(* Logix 5000 project; controller TFF vendor 1 type 14 code 107 rev 33.11; software revision 33.04; part 28 of 38 *)
(* tags used below, declared in another part *)
   Address : DINT;   // Temp Address
   AO1 : ALIAS FOR AnalogOutput[8];
   AO2 : ALIAS FOR AnalogOutput[9];
   AO3 : ALIAS FOR AnalogOutput[10];
   AO4 : ALIAS FOR AnalogOutput[11];
   ControlLoop_FeedBagLevel : ALIAS FOR ControlLoop[2];
   ControlLoop_FeedBagLevelAlarm : ALIAS FOR AlarmDeviation[2];
   DF48MIX : ALIAS FOR DigitalPoint[26];
   DF48P001 : ALIAS FOR DigitalPoint[23];
   DF48P002 : ALIAS FOR DigitalPoint[24];
   DigitalOutput : BOOL[256];   // Digital Output Array these bits are sent to output cards.
   DigitalPoint : DigitalPoint[150];   // Digital Point Array
   DO1 : ALIAS FOR DigitalOutput[80];
   DO2 : ALIAS FOR DigitalOutput[81];
   DO3 : ALIAS FOR DigitalOutput[82];
   DO4 : ALIAS FOR DigitalOutput[83];
   DO5 : ALIAS FOR DigitalOutput[84];
   DO6 : ALIAS FOR DigitalOutput[85];
   DO7 : ALIAS FOR DigitalOutput[86];
   Drive : Drive[11];   // Drives Array
   Exchange_OUT : Exchange_OUT;   // Exchange Outputs
   FlowPath : FlowPath[64];   // Flow Path Array
   MIX101DF : ALIAS FOR DigitalPoint[28];
   Mixer : Mixer;   // Mixer config. structure
   Options : Options;   // Options List
   Phase0 : ALIAS FOR Phase[0];   // Phase 0
   PI401 : ALIAS FOR AnalogPoint[8];
   PipeAnimation : PipeAnimation;   // HMI Pipe Animation Array
   SIC001DF : ALIAS FOR DigitalPoint[16];
   SIC002 : ALIAS FOR Drive[2];
   SIC002DF : ALIAS FOR DigitalPoint[17];
   SIC004 : ALIAS FOR Drive[3];
   SysControl : SysControl;   // General system status and command
   Tank : TankManagement;   // Tank Management
   WI101 : ALIAS FOR AnalogPoint[15];
(* Process, continued *)

ROUTINE Drive_SIC002_Transfer   (* ladder *)
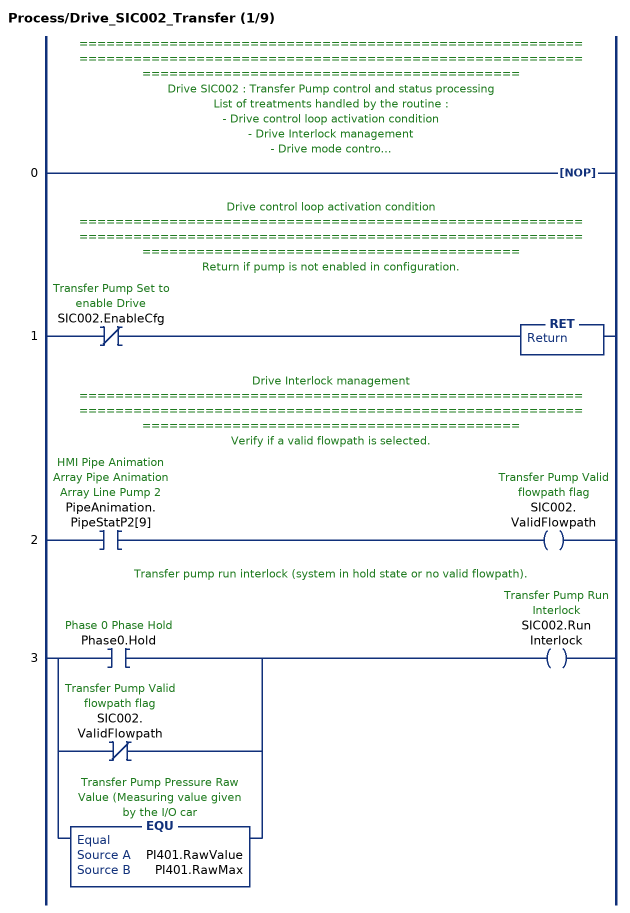
   // ==========================================================================================================================================================
   //                                                              Drive SIC002 : Transfer Pump control and status processing
   //                                                     List of treatments handled by the routine :
   //                                                          - Drive control loop activation condition
   //                                                          - Drive Interlock management
   //                                                          - Drive mode control
   //                                                          - Drive run command control
   //                                                          - Drive status management
   //                                                          - Drive status for HMI
   //                                                          - Drive DigitalOutput control
   //                                                     -----------------------------------------------------------------------------------------------------------------------------------------------------
   //                                                     History
   // 		2019-DEC-24 - Merck - Q. Spindler - Initial version for Candidate Release 1.00.00.00.a
   // 		2020-APR-06 - Merck - Q. Spindler - Modifications for Candidate Release 1.00.00.00.b
   //                                                                     - Add interlock when PI401 raw value is equal to RawMax (Sensor disconected)
   // ==========================================================================================================================================================
   0: NOP();
   // Drive control loop activation condition
   // ==========================================================================================================================================================
   // Return if pump is not enabled in configuration.
   1: XIO(SIC002.EnableCfg)RET();
   // Drive Interlock management
   // ==========================================================================================================================================================
   // Verify if a valid flowpath is selected.
   2: XIC(PipeAnimation.PipeStatP2[9])OTE(SIC002.ValidFlowpath);
   // Transfer pump run interlock (system in hold state or no valid flowpath).
   3: [XIC(Phase0.Hold) ,XIO(SIC002.ValidFlowpath) ,EQU(PI401.RawValue,PI401.RawMax) ]OTE(SIC002.RunInterlock);
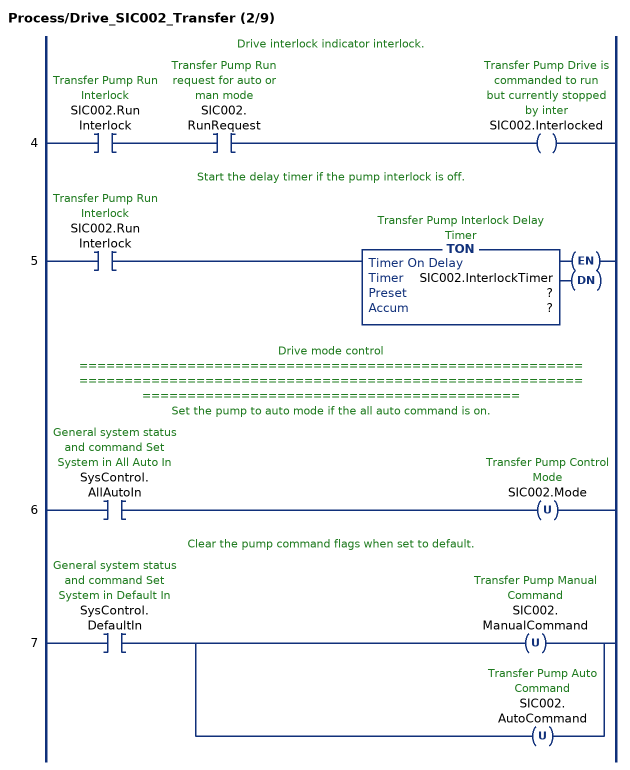
   // Drive interlock indicator interlock.
   4: XIC(SIC002.RunInterlock)XIC(SIC002.RunRequest)OTE(SIC002.Interlocked);
   // Start the delay timer if the pump interlock is off.
   5: XIC(SIC002.RunInterlock)TON(SIC002.InterlockTimer,?,?);
   // Drive mode control
   // ==========================================================================================================================================================
   // Set the pump to auto mode if the all auto command is on.
   6: XIC(SysControl.AllAutoIn)OTU(SIC002.Mode);
   // Clear the pump command flags when set to default.
   7: XIC(SysControl.DefaultIn)[OTU(SIC002.ManualCommand) ,OTU(SIC002.AutoCommand) ];
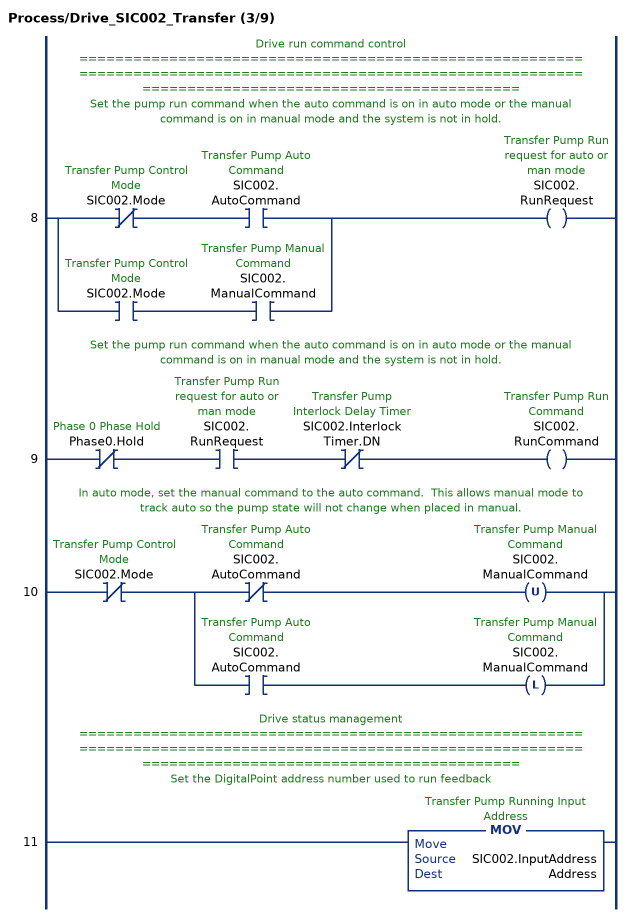
   // Drive run command control
   // ==========================================================================================================================================================
   // Set the pump run command when the auto command is on in auto mode or the manual command is on in manual mode and the system is not in hold.
   8: [XIO(SIC002.Mode) XIC(SIC002.AutoCommand) ,XIC(SIC002.Mode) XIC(SIC002.ManualCommand) ]OTE(SIC002.RunRequest);
   // Set the pump run command when the auto command is on in auto mode or the manual command is on in manual mode and the system is not in hold.
   9: XIO(Phase0.Hold)XIC(SIC002.RunRequest)XIO(SIC002.InterlockTimer.DN)OTE(SIC002.RunCommand);
   // In auto mode, set the manual command to the auto command.  This allows manual mode to track auto so the pump state will not change when placed in manual.
   10: XIO(SIC002.Mode)[XIO(SIC002.AutoCommand) OTU(SIC002.ManualCommand) ,XIC(SIC002.AutoCommand) OTL(SIC002.ManualCommand) ];
   // Drive status management
   // ==========================================================================================================================================================
   // Set the DigitalPoint address number used to run feedback
   11: MOV(SIC002.InputAddress,Address);
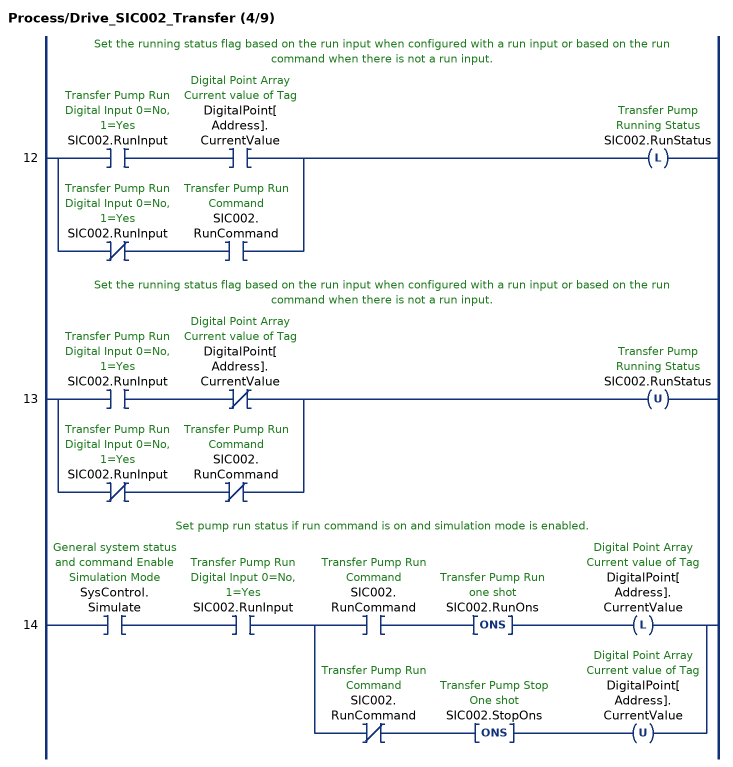
   // Set the running status flag based on the run input when configured with a run input or based on the run command when there is not a run input.
   12: [XIC(SIC002.RunInput) XIC(DigitalPoint[Address].CurrentValue) ,XIO(SIC002.RunInput) XIC(SIC002.RunCommand) ]OTL(SIC002.RunStatus);
   // Set the running status flag based on the run input when configured with a run input or based on the run command when there is not a run input.
   13: [XIC(SIC002.RunInput) XIO(DigitalPoint[Address].CurrentValue) ,XIO(SIC002.RunInput) XIO(SIC002.RunCommand) ]OTU(SIC002.RunStatus);
   // Set pump run status if run command is on and simulation mode is enabled.
   14: XIC(SysControl.Simulate)XIC(SIC002.RunInput)[XIC(SIC002.RunCommand) ONS(SIC002.RunOns) OTL(DigitalPoint[Address].CurrentValue) ,XIO(SIC002.RunCommand) ONS(SIC002.StopOns) OTU(DigitalPoint[Address].CurrentValue) ];
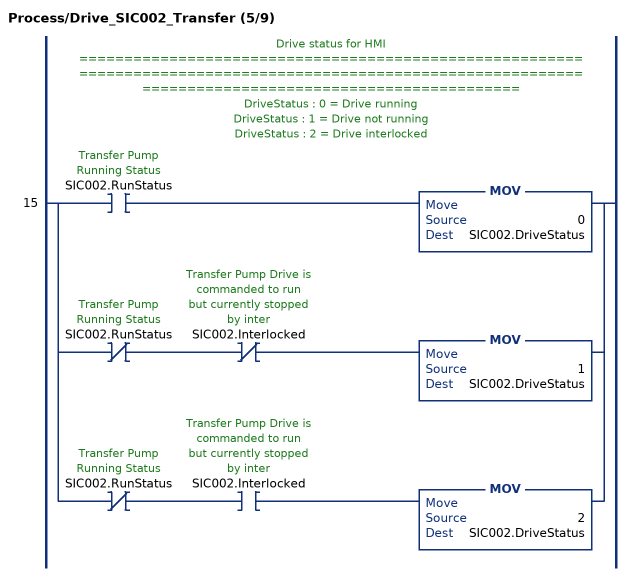
   // Drive status for HMI
   // ==========================================================================================================================================================
   //  DriveStatus : 0 = Drive running
   //  DriveStatus : 1 = Drive not running
   //  DriveStatus : 2 = Drive interlocked
   15: [XIC(SIC002.RunStatus) MOV(0,SIC002.DriveStatus) ,XIO(SIC002.RunStatus) XIO(SIC002.Interlocked) MOV(1,SIC002.DriveStatus) ,XIO(SIC002.RunStatus) XIC(SIC002.Interlocked) MOV(2,SIC002.DriveStatus) ];
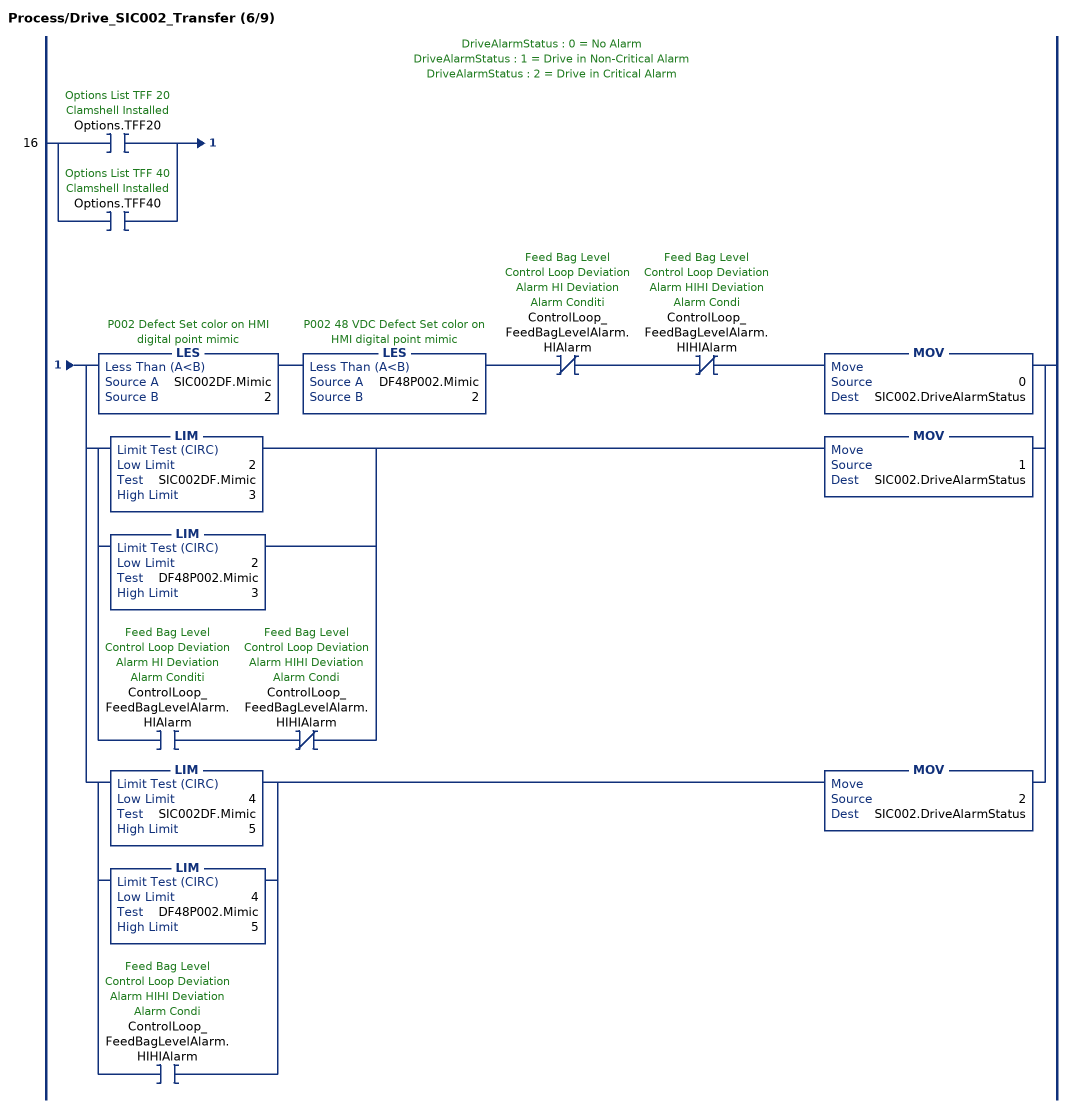
   // DriveAlarmStatus : 0 = No Alarm
   //  DriveAlarmStatus : 1 = Drive in Non-Critical Alarm
   //  DriveAlarmStatus : 2 = Drive in Critical Alarm
   16: [XIC(Options.TFF20) ,XIC(Options.TFF40) ][LES(SIC002DF.Mimic,2) LES(DF48P002.Mimic,2) XIO(ControlLoop_FeedBagLevelAlarm.HIAlarm) XIO(ControlLoop_FeedBagLevelAlarm.HIHIAlarm) MOV(0,SIC002.DriveAlarmStatus) ,[LIM(2,SIC002DF.Mimic,3) ,LIM(2,DF48P002.Mimic,3) ,XIC(ControlLoop_FeedBagLevelAlarm.HIAlarm) XIO(ControlLoop_FeedBagLevelAlarm.HIHIAlarm) ] MOV(1,SIC002.DriveAlarmStatus) ,[LIM(4,SIC002DF.Mimic,5) ,LIM(4,DF48P002.Mimic,5) ,XIC(ControlLoop_FeedBagLevelAlarm.HIHIAlarm) ] MOV(2,SIC002.DriveAlarmStatus) ];
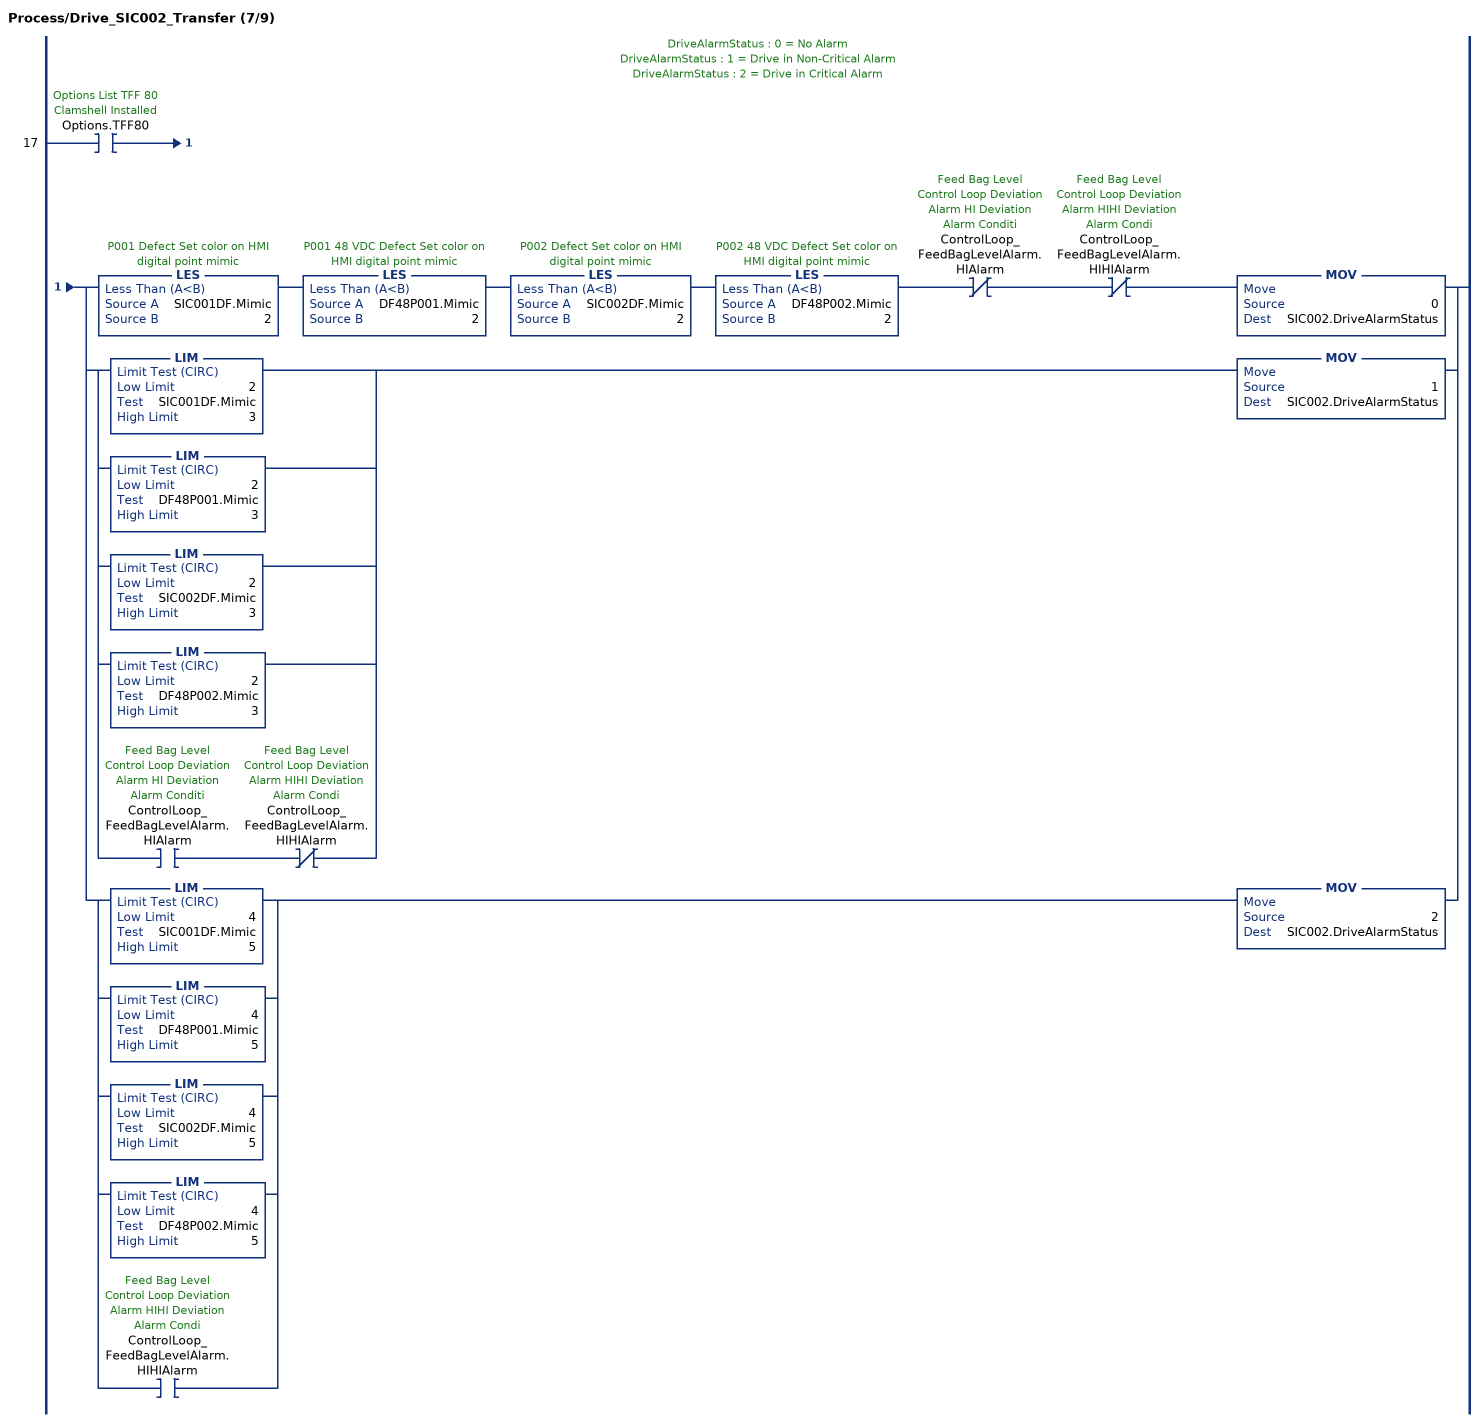
   // DriveAlarmStatus : 0 = No Alarm
   //  DriveAlarmStatus : 1 = Drive in Non-Critical Alarm
   //  DriveAlarmStatus : 2 = Drive in Critical Alarm
   17: XIC(Options.TFF80)[LES(SIC001DF.Mimic,2) LES(DF48P001.Mimic,2) LES(SIC002DF.Mimic,2) LES(DF48P002.Mimic,2) XIO(ControlLoop_FeedBagLevelAlarm.HIAlarm) XIO(ControlLoop_FeedBagLevelAlarm.HIHIAlarm) MOV(0,SIC002.DriveAlarmStatus) ,[LIM(2,SIC001DF.Mimic,3) ,LIM(2,DF48P001.Mimic,3) ,LIM(2,SIC002DF.Mimic,3) ,LIM(2,DF48P002.Mimic,3) ,XIC(ControlLoop_FeedBagLevelAlarm.HIAlarm) XIO(ControlLoop_FeedBagLevelAlarm.HIHIAlarm) ] MOV(1,SIC002.DriveAlarmStatus) ,[LIM(4,SIC001DF.Mimic,5) ,LIM(4,DF48P001.Mimic,5) ,LIM(4,SIC002DF.Mimic,5) ,LIM(4,DF48P002.Mimic,5) ,XIC(ControlLoop_FeedBagLevelAlarm.HIHIAlarm) ] MOV(2,SIC002.DriveAlarmStatus) ];
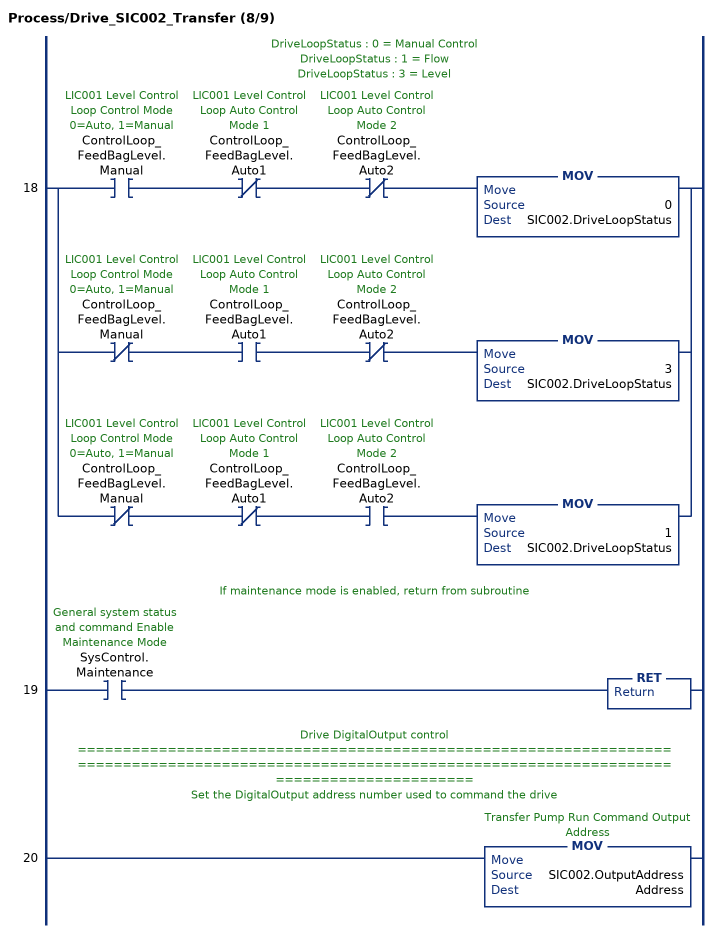
   // DriveLoopStatus : 0 = Manual Control
   //  DriveLoopStatus : 1 = Flow
   //  DriveLoopStatus : 3 = Level
   18: [XIC(ControlLoop_FeedBagLevel.Manual) XIO(ControlLoop_FeedBagLevel.Auto1) XIO(ControlLoop_FeedBagLevel.Auto2) MOV(0,SIC002.DriveLoopStatus) ,XIO(ControlLoop_FeedBagLevel.Manual) XIC(ControlLoop_FeedBagLevel.Auto1) XIO(ControlLoop_FeedBagLevel.Auto2) MOV(3,SIC002.DriveLoopStatus) ,XIO(ControlLoop_FeedBagLevel.Manual) XIO(ControlLoop_FeedBagLevel.Auto1) XIC(ControlLoop_FeedBagLevel.Auto2) MOV(1,SIC002.DriveLoopStatus) ];
   // If maintenance mode is enabled, return from subroutine
   19: XIC(SysControl.Maintenance)RET();
   // Drive DigitalOutput control
   // ==========================================================================================================================================================
   // Set the DigitalOutput address number used to command the drive
   20: MOV(SIC002.OutputAddress,Address);
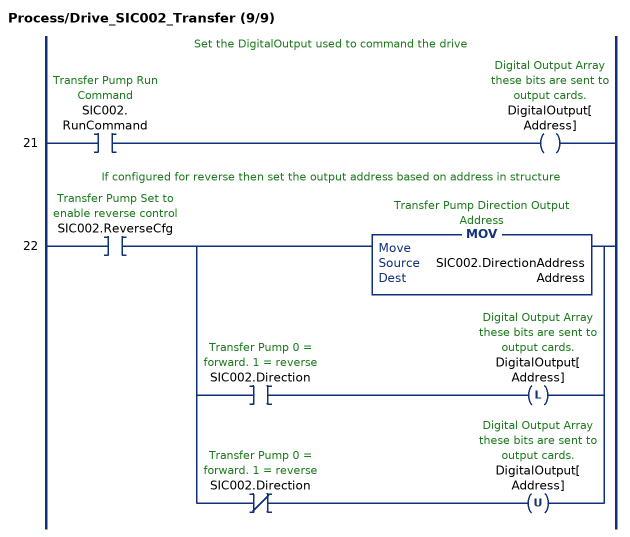
   // Set the DigitalOutput used to command the drive
   21: XIC(SIC002.RunCommand)OTE(DigitalOutput[Address]);
   // If configured for reverse then set the output address based on address in structure
   22: XIC(SIC002.ReverseCfg)[MOV(SIC002.DirectionAddress,Address) ,XIC(SIC002.Direction) OTL(DigitalOutput[Address]) ,XIO(SIC002.Direction) OTU(DigitalOutput[Address]) ];
END_ROUTINE

ROUTINE Drive_SIC004_Mixer   (* ladder *)
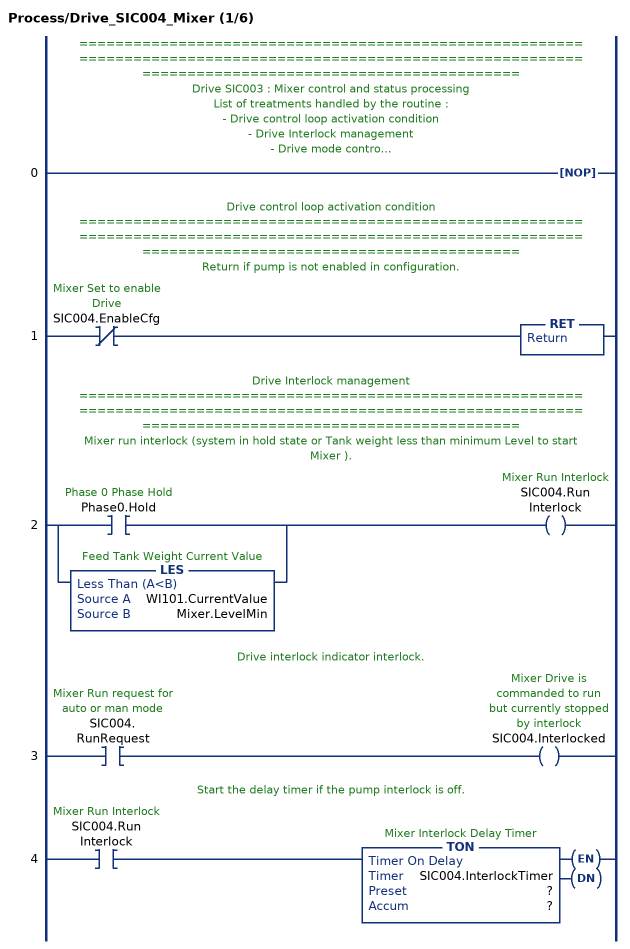
   // ==========================================================================================================================================================
   //                                                        Drive SIC003 : Mixer control and status processing
   //                                                     List of treatments handled by the routine :
   //                                                          - Drive control loop activation condition
   //                                                          - Drive Interlock management
   //                                                          - Drive mode control
   //                                                          - Drive run command control
   //                                                          - Drive status management
   //                                                          - Drive status for HMI
   //                                                          - Drive DigitalOutput control
   //                                                     -----------------------------------------------------------------------------------------------------------------------------------------------------
   //                                                     History
   // 		2019-DEC-24 - Merck - Q. Spindler - Initial version for Candidate Release 1.00.00.00.a
   // ==========================================================================================================================================================
   0: NOP();
   // Drive control loop activation condition
   // ==========================================================================================================================================================
   // Return if pump is not enabled in configuration.
   1: XIO(SIC004.EnableCfg)RET();
   // Drive Interlock management
   // ==========================================================================================================================================================
   // Mixer run interlock (system in hold state or Tank weight less than minimum Level to start Mixer ).
   2: [XIC(Phase0.Hold) ,LES(WI101.CurrentValue,Mixer.LevelMin) ]OTE(SIC004.RunInterlock);
   // Drive interlock indicator interlock.
   3: XIC(SIC004.RunRequest)OTE(SIC004.Interlocked);
   // Start the delay timer if the pump interlock is off.
   4: XIC(SIC004.RunInterlock)TON(SIC004.InterlockTimer,?,?);
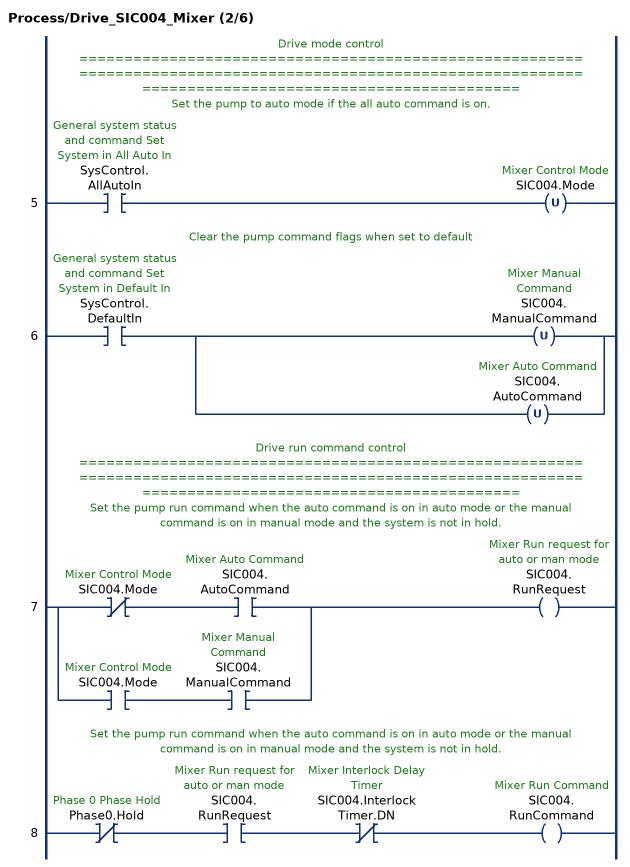
   // Drive mode control
   // ==========================================================================================================================================================
   // Set the pump to auto mode if the all auto command is on.
   5: XIC(SysControl.AllAutoIn)OTU(SIC004.Mode);
   // Clear the pump command flags when set to default
   6: XIC(SysControl.DefaultIn)[OTU(SIC004.ManualCommand) ,OTU(SIC004.AutoCommand) ];
   // Drive run command control
   // ==========================================================================================================================================================
   // Set the pump run command when the auto command is on in auto mode or the manual command is on in manual mode and the system is not in hold.
   7: [XIO(SIC004.Mode) XIC(SIC004.AutoCommand) ,XIC(SIC004.Mode) XIC(SIC004.ManualCommand) ]OTE(SIC004.RunRequest);
   // Set the pump run command when the auto command is on in auto mode or the manual command is on in manual mode and the system is not in hold.
   8: XIO(Phase0.Hold)XIC(SIC004.RunRequest)XIO(SIC004.InterlockTimer.DN)OTE(SIC004.RunCommand);
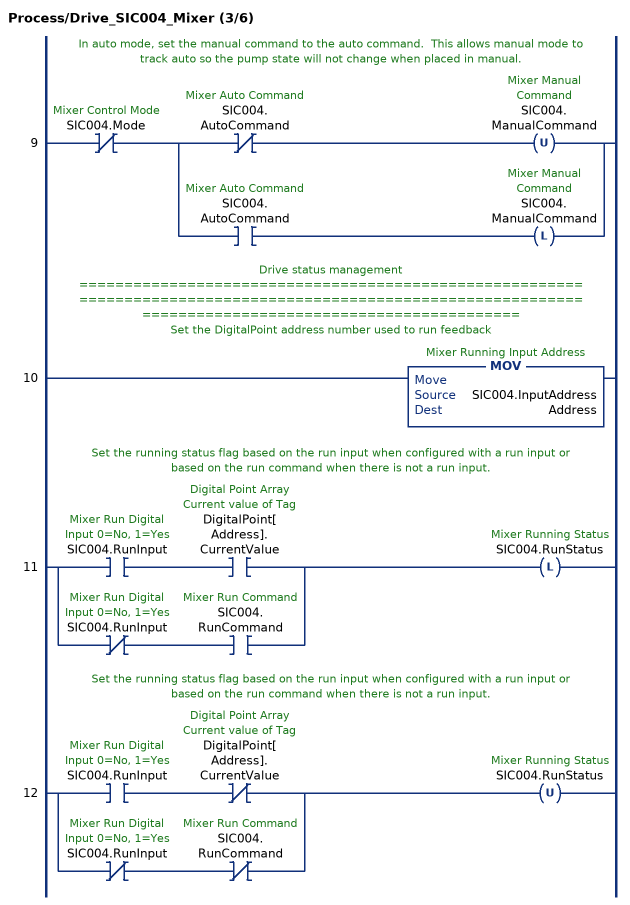
   // In auto mode, set the manual command to the auto command.  This allows manual mode to track auto so the pump state will not change when placed in manual.
   9: XIO(SIC004.Mode)[XIO(SIC004.AutoCommand) OTU(SIC004.ManualCommand) ,XIC(SIC004.AutoCommand) OTL(SIC004.ManualCommand) ];
   // Drive status management
   // ==========================================================================================================================================================
   // Set the DigitalPoint address number used to run feedback
   10: MOV(SIC004.InputAddress,Address);
   // Set the running status flag based on the run input when configured with a run input or based on the run command when there is not a run input.
   11: [XIC(SIC004.RunInput) XIC(DigitalPoint[Address].CurrentValue) ,XIO(SIC004.RunInput) XIC(SIC004.RunCommand) ]OTL(SIC004.RunStatus);
   // Set the running status flag based on the run input when configured with a run input or based on the run command when there is not a run input.
   12: [XIC(SIC004.RunInput) XIO(DigitalPoint[Address].CurrentValue) ,XIO(SIC004.RunInput) XIO(SIC004.RunCommand) ]OTU(SIC004.RunStatus);
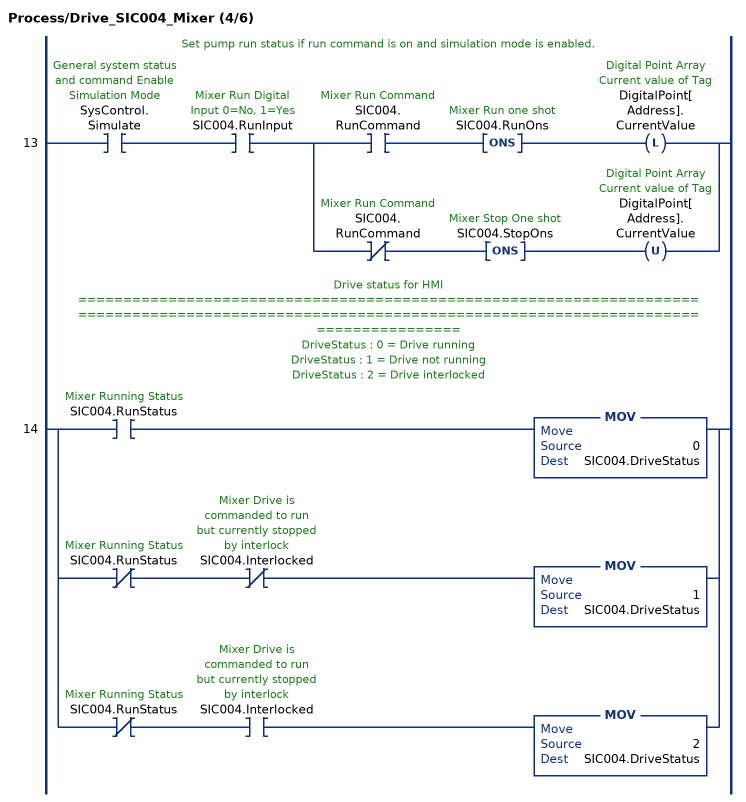
   // Set pump run status if run command is on and simulation mode is enabled.
   13: XIC(SysControl.Simulate)XIC(SIC004.RunInput)[XIC(SIC004.RunCommand) ONS(SIC004.RunOns) OTL(DigitalPoint[Address].CurrentValue) ,XIO(SIC004.RunCommand) ONS(SIC004.StopOns) OTU(DigitalPoint[Address].CurrentValue) ];
   // Drive status for HMI
   // ==========================================================================================================================================================
   //  DriveStatus : 0 = Drive running
   //  DriveStatus : 1 = Drive not running
   //  DriveStatus : 2 = Drive interlocked
   14: [XIC(SIC004.RunStatus) MOV(0,SIC004.DriveStatus) ,XIO(SIC004.RunStatus) XIO(SIC004.Interlocked) MOV(1,SIC004.DriveStatus) ,XIO(SIC004.RunStatus) XIC(SIC004.Interlocked) MOV(2,SIC004.DriveStatus) ];
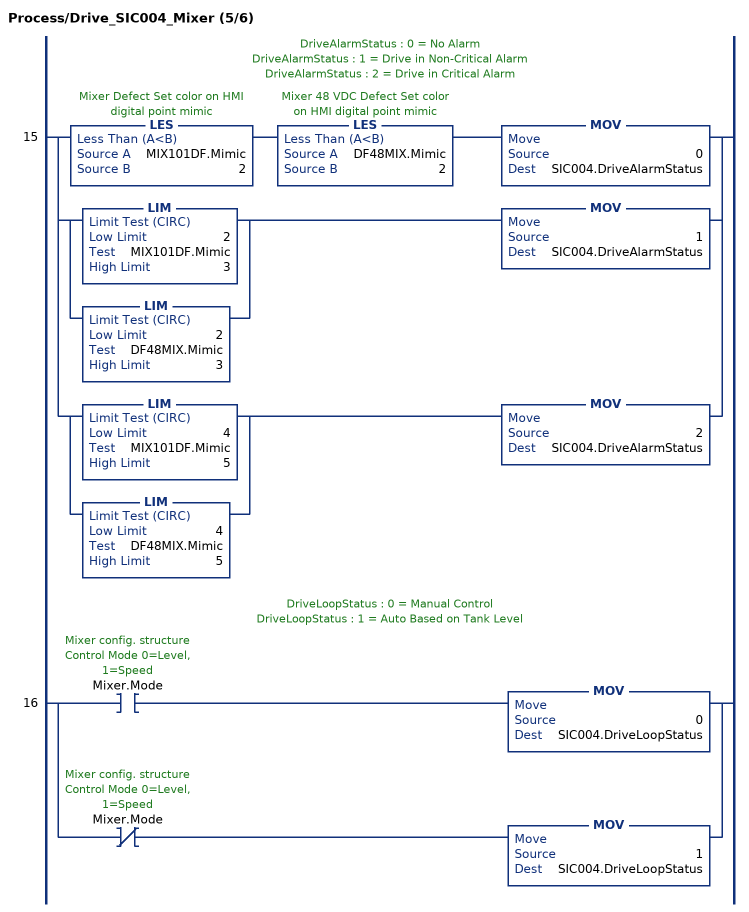
   // DriveAlarmStatus : 0 = No Alarm
   //  DriveAlarmStatus : 1 = Drive in Non-Critical Alarm
   //  DriveAlarmStatus : 2 = Drive in Critical Alarm
   15: [LES(MIX101DF.Mimic,2) LES(DF48MIX.Mimic,2) MOV(0,SIC004.DriveAlarmStatus) ,[LIM(2,MIX101DF.Mimic,3) ,LIM(2,DF48MIX.Mimic,3) ] MOV(1,SIC004.DriveAlarmStatus) ,[LIM(4,MIX101DF.Mimic,5) ,LIM(4,DF48MIX.Mimic,5) ] MOV(2,SIC004.DriveAlarmStatus) ];
   // DriveLoopStatus : 0 = Manual Control
   //  DriveLoopStatus : 1 = Auto Based on Tank Level
   16: [XIC(Mixer.Mode) MOV(0,SIC004.DriveLoopStatus) ,XIO(Mixer.Mode) MOV(1,SIC004.DriveLoopStatus) ];
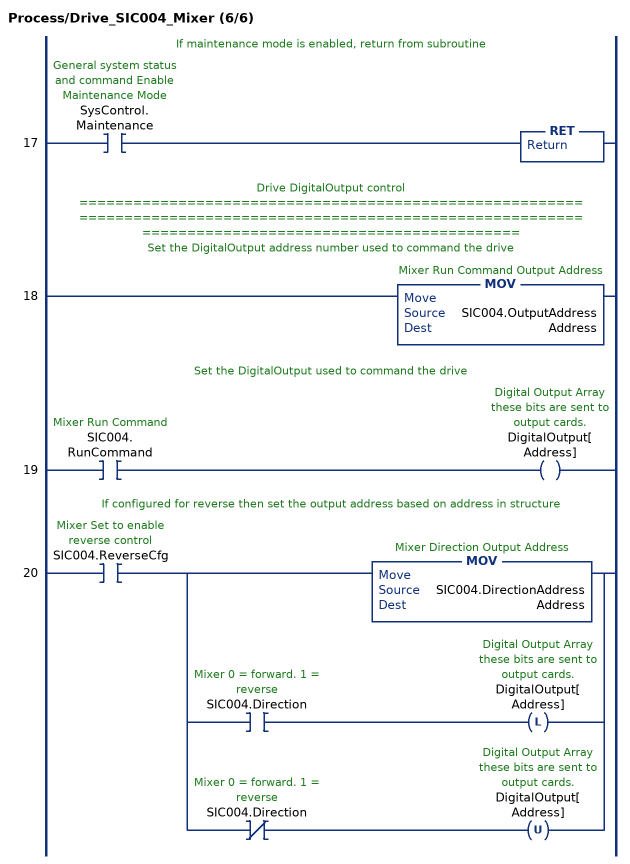
   // If maintenance mode is enabled, return from subroutine
   17: XIC(SysControl.Maintenance)RET();
   // Drive DigitalOutput control
   // ==========================================================================================================================================================
   // Set the DigitalOutput address number used to command the drive
   18: MOV(SIC004.OutputAddress,Address);
   // Set the DigitalOutput used to command the drive
   19: XIC(SIC004.RunCommand)OTE(DigitalOutput[Address]);
   // If configured for reverse then set the output address based on address in structure
   20: XIC(SIC004.ReverseCfg)[MOV(SIC004.DirectionAddress,Address) ,XIC(SIC004.Direction) OTL(DigitalOutput[Address]) ,XIO(SIC004.Direction) OTU(DigitalOutput[Address]) ];
END_ROUTINE

ROUTINE Drives   (* ladder *)
// Pump Control Routine
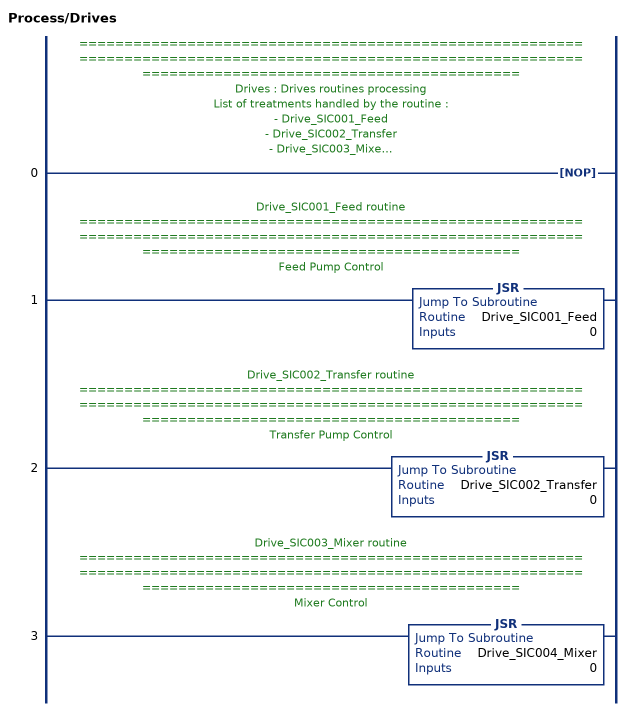
   // ==========================================================================================================================================================
   //                                                                                                                           Drives : Drives routines processing
   //                                                     List of treatments handled by the routine :
   //                                                          - Drive_SIC001_Feed
   //                                                          - Drive_SIC002_Transfer
   //                                                          - Drive_SIC003_Mixer
   //                                                     -----------------------------------------------------------------------------------------------------------------------------------------------------
   //                                                     History
   // 		2019-DEC-24 - Merck - Q. Spindler - Initial version for Candidate Release 1.00.00.00.a
   // ==========================================================================================================================================================
   0: NOP();
   // Drive_SIC001_Feed routine
   // ==========================================================================================================================================================
   // Feed Pump Control
   1: JSR(Drive_SIC001_Feed,0);
   // Drive_SIC002_Transfer routine
   // ==========================================================================================================================================================
   // Transfer Pump Control
   2: JSR(Drive_SIC002_Transfer,0);
   // Drive_SIC003_Mixer routine
   // ==========================================================================================================================================================
   // Mixer Control
   3: JSR(Drive_SIC004_Mixer,0);
END_ROUTINE

ROUTINE Exchange_IO   (* ladder *)
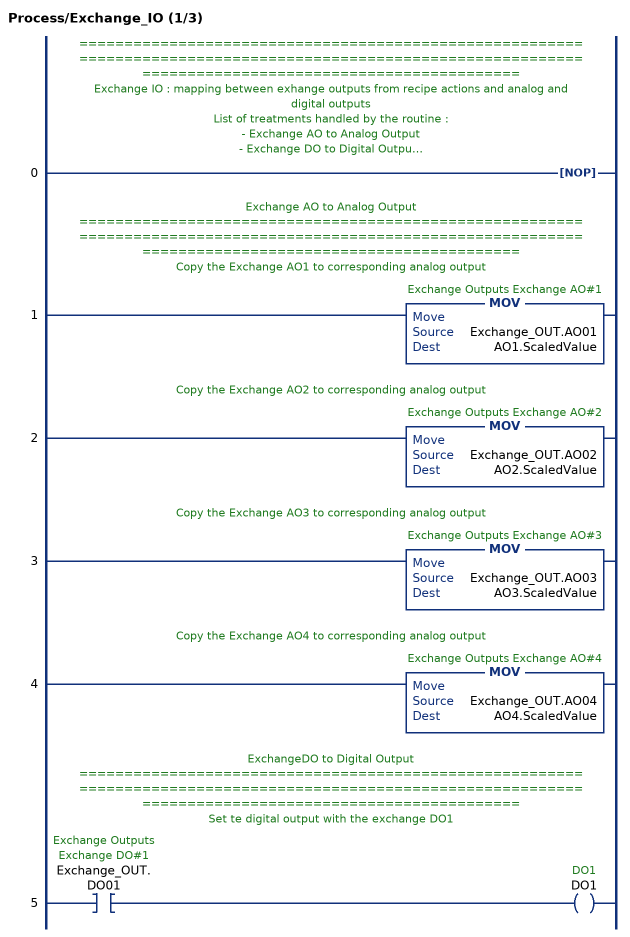
   // ==========================================================================================================================================================
   //                                                                             Exchange IO : mapping between exhange outputs from recipe actions and analog and digital outputs
   //                                                     List of treatments handled by the routine :
   //                                                          - Exchange AO to Analog Output
   //                                                          - Exchange DO to Digital Output
   //                                                     -----------------------------------------------------------------------------------------------------------------------------------------------------
   //                                                     History
   // 		2019-DEC-24 - Merck - Q. Spindler - Initial version for Candidate Release 1.00.00.00.a
   // ==========================================================================================================================================================
   0: NOP();
   // Exchange AO to Analog Output
   // ==========================================================================================================================================================
   // Copy the Exchange AO1 to corresponding analog output
   1: MOV(Exchange_OUT.AO01,AO1.ScaledValue);
   // Copy the Exchange AO2 to corresponding analog output
   2: MOV(Exchange_OUT.AO02,AO2.ScaledValue);
   // Copy the Exchange AO3 to corresponding analog output
   3: MOV(Exchange_OUT.AO03,AO3.ScaledValue);
   // Copy the Exchange AO4 to corresponding analog output
   4: MOV(Exchange_OUT.AO04,AO4.ScaledValue);
   // ExchangeDO to Digital Output
   // ==========================================================================================================================================================
   // Set te digital output with the exchange DO1
   5: XIC(Exchange_OUT.DO01)OTE(DO1);
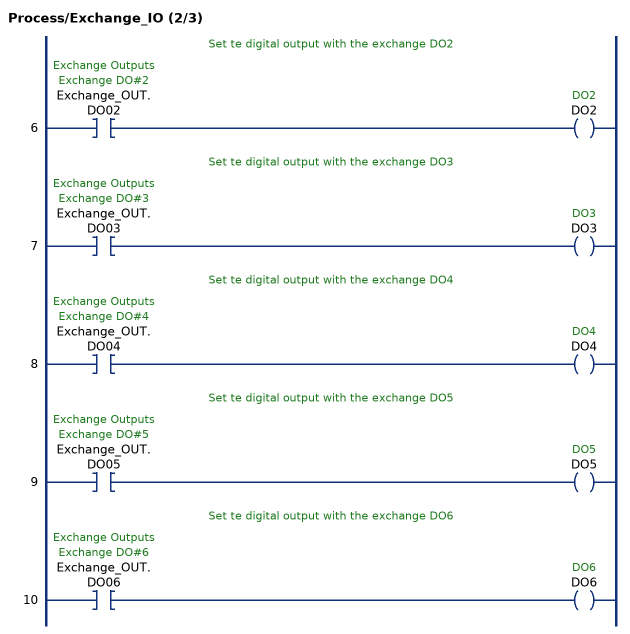
   // Set te digital output with the exchange DO2
   6: XIC(Exchange_OUT.DO02)OTE(DO2);
   // Set te digital output with the exchange DO3
   7: XIC(Exchange_OUT.DO03)OTE(DO3);
   // Set te digital output with the exchange DO4
   8: XIC(Exchange_OUT.DO04)OTE(DO4);
   // Set te digital output with the exchange DO5
   9: XIC(Exchange_OUT.DO05)OTE(DO5);
   // Set te digital output with the exchange DO6
   10: XIC(Exchange_OUT.DO06)OTE(DO6);
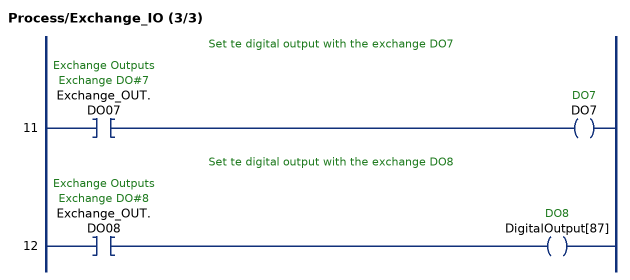
   // Set te digital output with the exchange DO7
   11: XIC(Exchange_OUT.DO07)OTE(DO7);
   // Set te digital output with the exchange DO8
   12: XIC(Exchange_OUT.DO08)OTE(DigitalOutput[87]);
END_ROUTINE
